(* IEC 61131-3 sources: rusty/tests/lit/multi/external_enum_variants, 3 files *)

(* ---- base.st ---- *)
TYPE Color : (Red, Green, Blue); END_TYPE

VAR_GLOBAL
    gColor : Color := Green;
END_VAR

(* ---- main.st ---- *)
FUNCTION main : DINT
VAR
    fb : ColorFb;
    c : Color;
END_VAR
    printf('%d$N', gColor);
    fb();
    printf('%d$N', fb.out);
    c := next_color(fb.out);
    printf('%d$N', c);
    CASE c OF
        Green: printf('green$N');
        ELSE printf('other$N');
    END_CASE
    gColor := Blue;
    printf('%d$N', gColor);
END_FUNCTION

(* ---- lib.st ---- *)
FUNCTION_BLOCK ColorFb
VAR_OUTPUT
    out : Color := Blue;
END_VAR
    IF gColor = Green THEN
        out := Red;
    END_IF
END_FUNCTION_BLOCK

FUNCTION next_color : Color
VAR_INPUT
    c : Color;
END_VAR
    CASE c OF
        Red: next_color := Green;
        Green: next_color := Blue;
        Blue: next_color := Red;
    END_CASE
END_FUNCTION
